Fanuc KAREL source: KO00097.KL

PROGRAM KO00097
%NOLOCKGROUP
VAR
  A: INTEGER
  B: INTEGER
  OUT: INTEGER
BEGIN
  A = 1
  B = 2
  OUT = ATAN2(A, B)
END KO00097
